TYPE ST_ParentChildControl :
STRUCT
	mode				: E_SystemMode;
	state				: INT;
	//sequencerState		: E_SequenceState;
	instancePath		: T_MaxString := '';
	
	estop				: BOOL;
END_STRUCT
END_TYPE

(* stored: Version 1.1.0.1, ProductVersion 3.1.4024.12
   DUT ST_ParentChildControl: Id {2c789bdd-4224-4a0c-a03a-ff017fa08b41} *)
